(* IEC 61131-3 sources: Masterarbeit/sigmatek/lasalclass2/PW022_hardware/Class/_DriveMngBase (part 2) *)

    for x := 0 to SDDMAXENTRIES -1 do
      if (AxBuffer[x].pThis <> NIL) then
        if(AxBuffer[x].InitFinished = FALSE) & (AxBuffer[x].AxisOk = 1) then
          return;
        end_if;
      else
        exit;
      end_if;
    end_for;

    bdSettings.AxisInit := TRUE;

    if bVaranConnected then
      toVaran.ExternInitFinished();
    else
      MyPara.uiCmd := BUSIF_DRIVEMNGBASE_EXTERN_INIT_FINISH;
      ToBusIF.NewInst(#MyPara, #MyResult);
    end_if;

END_FUNCTION

FUNCTION _DriveMngBase::ResetAxisInit
  VAR
  	x       : USINT;
  END_VAR

    for x := 0 to SDDMAXENTRIES -1 do
      if (AxBuffer[x].pThis <> NIL) then
        if (AxBuffer[x].AxisOk = 1) then
          AxBuffer[x].InitFinished := FALSE;
        end_if;
      end_if;
    end_for;

END_FUNCTION

FUNCTION GLOBAL _DriveMngBase::CommunicationState
	VAR_OUTPUT
		retcode 	: DINT;
	END_VAR

  retcode := cOnline;

END_FUNCTION

FUNCTION _DriveMngBase::L2CmdFinished
	VAR_INPUT
		pPara 	: ^CmdStruct;
		pResult 	: ^results;
	END_VAR
	VAR_OUTPUT
		ret_code 	: iprStates;
	END_VAR

  ret_code := READY;

  L2Buffer[L2WrIndex].AxisNo := to_usint(pPara^.aPara[3]);
  L2Buffer[L2WrIndex].ParRW := to_usint(pPara^.aPara[1]);
  L2Buffer[L2WrIndex].ParNo := to_usint(pPara^.aPara[0]);
  L2Buffer[L2WrIndex].ParValue := pPara^.aPara[2];
  L2Buffer[L2WrIndex].bActive := TRUE;

  if pPara^.uiCmd = SDD_ASYNC_READY then
    L2Buffer[L2WrIndex].ParState := 0;
  else
    L2Buffer[L2WrIndex].ParState := 1;
    L2Buffer[L2WrIndex].ParError := to_sint(pPara^.aPara[4]);
  end_if;

  L2WrIndex += 1;
  L2NewEntry += 1;
  if L2WrIndex > (L2MAXINDEX - 1) then
    L2WrIndex := 0;
  end_if;

END_FUNCTION

FUNCTION VIRTUAL GLOBAL _DriveMngBase::CmdState::NewInst
	VAR_INPUT
		pPara 	: ^CmdStruct;
		pResult 	: ^results;
	END_VAR
	VAR_OUTPUT
		ret_code 	: iprStates;
	END_VAR
  VAR
    AxisNo          : USINT;
    ParRW           : USINT;
    ParNo           : USINT;
    retcode         : DINT;
    AxIndex         : USINT;
    RetcodeSizeLeft : UDINT;
    pActRetEntry    : ^_ParaRefreshBufEntry;
    i               : USINT;
    pThisRes        : ^UDINT;
    FoundAxis       : USINT;

    // Variables for CMD_GET_HARDWARE_DIAGNOSIS and CMD_GET_HARDWARE_TREE_ENTRY
    pStr_HWTRequested         : ^CHAR;
    us_HWTRequestedCurrIndex  : USINT;
    us_RequestedPlace         : USINT;
    us_RequestedAxis          : USINT;
    us_NextAxis               : USINT;
    us_NextPlace              : USINT;
    ud_StrSize                : UDINT;
    ud_TempSerNo              : UDINT;

    MyPara   : CmdStruct;
    MyResult : results;
  END_VAR

  pStr_HWTRequested         := NIL;
  us_HWTRequestedCurrIndex  := 0;
  us_RequestedPlace         := 16#FF;
  us_RequestedAxis          := 16#FF;
  us_NextAxis               := 16#FF;
  us_NextPlace              := 16#FF;
  ud_StrSize                := 0;
  ud_TempSerNo              := 0;

  ret_code := READY;

  CASE pPara^.uiCmd OF
  SDD_ASYNC_READY :

    // check the parameter number
    case (pPara^.aPara[0]) of

    SDD_I_HW :

      HWVersion := pPara^.aPara[2];
      DriveType := GetDriveType(pPara^.aPara[2]);
      bdWait4HwInfoResponse.I_HW := FALSE;

    SDD_I_TYPE :

      Parameter_I_Type := pPara^.aPara[2];
      bdWait4HwInfoResponse.I_Type := FALSE;

    SDD_I_SER :

      SerialNo := pPara^.aPara[2];
      bdWait4HwInfoResponse.I_SER := FALSE;

    SDD_I_FW :

      FwVersionInt :=  pPara^.aPara[2];
      bdWait4HwInfoResponse.I_FW := FALSE;
      SetFWVersion();

    SDD_I_BUILD :

      FWDateInt :=  pPara^.aPara[2]$UDINT;
      bdWait4HwInfoResponse.I_BUILD := FALSE;
      SetFwDate();

    else

      // Parameter for log file are dependent on the drive, usParaLogIdx is set in GetLogFileCyclic
      if pPara^.aPara[0] = s_LogFileV.usParaLogIdx then
        s_LogFileV.dParaLogValRd     := pPara^.aPara[2];
        s_LogFileV.bWait4LogFilePara := FALSE;
      end_if;

    end_case;

  SDD_ASYNC_ERROR :
    case pPara^.aPara[0] of

    SDD_I_HW :

      HWVersion := 16#7FFFFFFF;
      DriveType := _NotFound;
      bdWait4HwInfoResponse.I_HW := FALSE;

    SDD_I_TYPE :

      Parameter_I_Type := 16#7FFFFFFF;
      bdWait4HwInfoResponse.I_Type := FALSE;

    SDD_I_SER :

      SerialNo := 16#7FFFFFFF;
      bdWait4HwInfoResponse.I_SER := FALSE;

    SDD_I_FW :

      FwVersionInt :=  16#7FFFFFFF;
      bdWait4HwInfoResponse.I_FW := FALSE;

    SDD_I_BUILD :

      FWDateInt :=  16#7FFFFFFF;
      bdWait4HwInfoResponse.I_BUILD := FALSE;

    else

      // Parameter for log file are dependent on the drive, usParaLogIdx is set in GetLogFileCyclic
      if pPara^.aPara[0] = s_LogFileV.usParaLogIdx then
        s_LogFileV.dParaLogValRd     := 16#7FFFFFFF;
        s_LogFileV.bWait4LogFilePara := FALSE;
      end_if;

    end_case;

  SDD_GETVERSION :
    ret_code := READY;
    pResult^.uiLng := sizeof(UINT);
    pResult^.aData[0] := SDD_L2VERSION;
    pResult^.aData[1] := 0;

  SDD_ONLINEOK :

    ret_code := READY;
    pResult^.uiLng := sizeof(USINT);
    pResult^.aData[0] := to_usint(Online.read());

    // if the ringbuffer is allocated
    if ChangesRingBuffer.pStart then
      // we reset the ringbuffer which contains the changes
      ChangesRingBuffer.ActEntries := 0;
      ChangesRingBuffer.pWrite := ChangesRingBuffer.pRead := ChangesRingBuffer.pStart;
      _memset(ChangesRingBuffer.pStart, 16#00, SDDBUFFERENTRY*sizeof(_ParaRefreshBufEntry));
    end_if;

  SDD_RWPARLASAL2 :

    if Online.read() = 1 then
      ret_code := BUSY;

      // get Axisnumber
      AxisNo := to_usint(pPara^.aPara[0] AND 16#FF);

      // on SDD210 or SDD215 we fake the axis number of the 2nd axis for external use, so we have to correct it here
      if b_IsSDD21x & (AxisNo = 2) then // RamAnd 22.09.2010 16:12
        AxisNo := 3;
      end_if;

      AxIndex := GetAxIndex(AxisNo-1);

      if AxIndex = 16#FF then
        ret_code := ERROR;
        return;
      end_if;

      // read or write
      ParRw   := to_usint((pPara^.aPara[0] AND 16#FF00) SHR 8);
      // parameter number
      ParNo   := to_usint((pPara^.aPara[0] AND 16#FF0000) SHR 16);

      case ParRw of
      0 : // Read the parameter
        //if right I-HC code and scope buffer request then read 12 byte drive scope data over ID 0x2080 and SubID 0x09 is allowed
        if ((HWVersion and DRIVEMNG_DRIVESCOPE_SCOPE_BIT) = DRIVEMNG_DRIVESCOPE_SCOPE_BIT)
        & bLasalErrorBufferRequest = FALSE then

          case ParNo of
            251:
              AddASyncEntryDS402(AxisNo:=AxIndex, uiParaID:=DRIVEMNG_DRIVESCOPE_GETALL_PARAM, usParaSubID:=9, usRdWr:=0, pValue:=Nil, bsDataInfo:=2, pThisObj:= this, usEntry:=3);
              ret_code := Busy;

            252:
              //use always zero for SDD1X00 scope data
              pPara^.aPara[0] := (pPara^.aPara[0] AND (16#FFFFFF00)$DINT);
              ret_code := CmdState.GetState(pPara:=pPara, pResult:=pResult);

            253:
              //use always zero for SDD1X00 scope data
              pPara^.aPara[0] := (pPara^.aPara[0] AND (16#FFFFFF00)$DINT);
              ret_code := CmdState.GetState(pPara:=pPara, pResult:=pResult);

          else
            retcode := AddASyncEntry(AxisNo:= AxIndex, usParaNr:= ParNo , usRdWr:= ParRw, dValue:=0, pThisObj:= this, usEntry:=3);
          end_case;
        else
          retcode := AddASyncEntry(AxisNo:= AxIndex, usParaNr:= ParNo , usRdWr:= ParRw, dValue:=0, pThisObj:= this, usEntry:=3);
        end_if;

      1 : // Write the parameter
        //if right I-HC code then read 12 byte drive scope data over ID 0x2080 and SubID 0x09 is allowed
        if ((HWVersion and DRIVEMNG_DRIVESCOPE_SCOPE_BIT) = DRIVEMNG_DRIVESCOPE_SCOPE_BIT) then
          if ParNo = 249 then
            //remember which request come from Lasal2 (Drive Scope or Errorbuffer)
            if pPara^.aPara[1] > DRIVEMNG_DRIVESCOPE_SINDEX_RANGE then
              bLasalErrorBufferRequest := TRUE;
            else
              bLasalErrorBufferRequest := FALSE;
            end_if;
          end_if;
        end_if;

        retcode := AddASyncEntry(AxisNo:= AxIndex, usParaNr:= ParNo , usRdWr:= ParRw, dValue:=pPara^.aPara[1], pThisObj:= this, usEntry:=3);
      else
        ret_code := ERROR;
      end_case;

      if retcode < 0 then
        // internal failure
        Ret_code := ERROR;
      end_if;
    else
      ret_code := ERROR;
    end_if;

  SDD_GETAXISINUSE :
    ret_code := READY;
    pResult^.uiLng := sizeof(BDINT);
    pResult^.aData[0]$BDINT :=  AxIndizesL2;

  SDD_GETSERIE :
    retcode := READY;
    pResult^.uiLng := sizeof(USINT);
    if bVaranConnected then
      pResult^.aData[0] := toVaran.GetSeries();
    else
      //sdias drive connected
      MyPara.uiCmd  := BUSIF_DRIVEMNGBASE_SDD_GETSERIES;
      ToBusIF.NewInst(#MyPara, #MyResult);
      pResult^.aData[0] := MyResult.aData[0];
    end_if;

  // new commands in lasal communication version 4 (SDD_GET_CHANGE_CNT, SDD_GET_PARAMS)
  SDD_GET_CHANGE_CNT :
    retcode := READY;
    pResult^.uiLng := sizeof(UDINT);
    pResult^.aData[0]$^DINT := #ChangesRingBuffer.ActEntries;

  SDD_GET_PARAMS :
    retcode := READY;
    if ChangesRingBuffer.ActEntries then

      RetcodeSizeLeft := sizeof(pResult^.aData) - SIZEOF(UINT);
      pResult^.uiLng := 0;

      pActRetEntry := (#pResult^.aData[2])$^_ParaRefreshBufEntry;

      // as long as there are entries in change buffer and we still have some place in the return value array
      while ChangesRingBuffer.ActEntries & (RetcodeSizeLeft > sizeof(_ParaRefreshBufEntry)) do

        // store actual buffer entry in returncode
        pActRetEntry^ := ChangesRingBuffer.pRead^;

        // increase size of returncode in it's header
        pResult^.uiLng += sizeof(_ParaRefreshBufEntry);

        // decrease available size of returncode
        RetcodeSizeLeft -= sizeof(_ParaRefreshBufEntry);

        // increase pointer in retcode
        pActRetEntry += sizeof(_ParaRefreshBufEntry);

        // increase read pointer in ring buffer
        ChangesRingBuffer.pRead += sizeof(_ParaRefreshBufEntry);
        if ChangesRingBuffer.pRead >= ChangesRingBuffer.pEnd then
          ChangesRingBuffer.pRead := ChangesRingBuffer.pStart;
        end_if;

        // decrease available changes
        ChangesRingBuffer.ActEntries -= 1;
      end_while;

      // save number of entries in the first 2 byte of the array
      pResult^.aData[0]$UINT := pResult^.uiLng / sizeof(_ParaRefreshBufEntry);

      LastRetcode := pResult^;
    else
      // no changes to fetch
      pResult^.uiLng := 0;
    end_if;

  //++++++++++++++++++++++++++++++++++++++++++++++++++++++++++++++++++++++++++++++++++++++++++++++++++++++++++++++++++++
  SDD_GET_AXIS_PTR_LIST:

    ret_code := READY;

    //                    NoAxis    +  Thisptr per axis
    pResult^.uiLng := (sizeof(DINT) + AxCount * sizeof(UDINT))$UINT;

    // get no of axis
    pResult^.aData[0]$DINT := AxCount;

    // get this pointer of axis to resultbuffer (with increasing AxNumber)
    pThisRes := #pResult^.aData[4]$UDINT;
    FoundAxis := 0;
    for i := 0 to SDDMAXENTRIES-1 do
      AxIndex := GetAxIndexByAxisBit(1 SHL i);
      if AxIndex <> 16#FF then
        FoundAxis += 1;
        pThisRes^ := AxBuffer[AxIndex].pThis$UDINT;
        pThisRes += sizeof(UDINT);
      end_if;
      if FoundAxis = AxCount then
        // all avaliable found, exit loop
        exit;
      end_if;
    end_for;
    // fill space with NIL if a axis is not found
    while FoundAxis < AxCount do
      pThisRes^ := NIL;
      pThisRes += sizeof(UDINT);
      FoundAxis += 1;
    end_while;

  //++++++++++++++++++++++++++++++++++++++++++++++++++++++++++++++++++++++++++++++++++++++++++++++++++++++++++++++++++++
  CMD_GET_HARDWARE_DIAGNOSIS :

    pResult^.aData$t_HWCGetHardwareDiagnosisOut.retcode := _HWC_RETVAL_ERROR;
    ret_code := ERROR;

    pStr_HWTRequested := pPara^.aPara[0]$t_HWCGetHardwareDiagnosisIn.pStr_HardewareTreeEntry;

    // Check HWT String
    if pStr_HWTRequested then

      us_HWTRequestedCurrIndex := to_usint(pStr_HWTRequested$^UINT^ + 1); // +1 for 2byte length, points to end of HWT String

      if ( (pStr_HWTRequested + us_HWTRequestedCurrIndex - 1)^ = HWT_ESCAPE_DRIVE ) then // second to last byte is Drive escape sequence

        us_RequestedPlace := (pStr_HWTRequested + us_HWTRequestedCurrIndex)^; // Get passed place

        // Return State and Device ID and set retcode ----------------------------------------------------------
        pResult^.aData$t_HWCGetHardwareDiagnosisOut.ClassState := CmdState;

        pResult^.aData$t_HWCGetHardwareDiagnosisOut.ud_DeviceID := GetDrvDeviceID();

        if CmdState = _NoHardware then
          pResult^.aData$t_HWCGetHardwareDiagnosisOut.retcode := _HWC_RETVAL_ERROR_NO_HARDWARE;
        elsif CmdState = _WrongHardware then
          pResult^.aData$t_HWCGetHardwareDiagnosisOut.retcode := _HWC_RETVAL_ERROR_WRONG_HARDWARE;
        elsif CmdState = _NoCalibDataFound then
          pResult^.aData$t_HWCGetHardwareDiagnosisOut.retcode := _HWC_RETVAL_ERROR_NO_CALIB_DATA_FOUND;
        elsif CmdState <> _ClassOk then
          pResult^.aData$t_HWCGetHardwareDiagnosisOut.retcode := _HWC_RETVAL_ERROR_NO_HARDWARE;
        end_if;
        //------------------------------------------------------------------------------------------------------

        if CmdState= _ClassOk then

          // Search for Axis with the passed place
          for i := 0 to SDDMAXENTRIES - 1 do
            if AxBuffer[i].pThis then

              if ( AxBuffer[i].Place  = us_RequestedPlace ) then

                // Diagnosis info is stored with the axis class
                ret_code := AxBuffer[i].pThis$pVirtualBase^.NewInst(pPara, pResult);

                // FW Version ----------------------------------------------------------------------------------------------------------
                pResult^.aData[0]$t_HWCGetHardwareDiagnosisOut.pStr_FWVersion := #a_FWVersion[0];  // Will be overwritten if this pointer is not equal

                ud_StrSize := FwNumStr.GetLength() ;
                pResult^.aData[0]$t_HWCGetHardwareDiagnosisOut.pStr_FWVersion     := NIL;

                if ud_StrSize then

                  if (ud_StrSize < sizeof(a_FWVersion)) then // < to account for 0 termination
                    // Copy complete string
                    FwNumStr.GetDataAt(pData:=#a_FWVersion[0], udSize:=ud_StrSize, udAt:=0);
                    a_FWVersion[ud_StrSize] := 0; // 0 termination
                  else
                    // Copy part string
                    FwNumStr.GetDataAt(pData:=#a_FWVersion[0], udSize:=sizeof(a_FWVersion)-1, udAt:=0);
                    a_FWVersion[sizeof(a_FWVersion)-1] := 0; // 0 termination
                  end_if;

                  pResult^.aData[0]$t_HWCGetHardwareDiagnosisOut.pStr_FWVersion := #a_FWVersion[0];
                end_if;

                // HW Version
                pResult^.aData[0]$t_HWCGetHardwareDiagnosisOut.hd_HWVersion := HWVersion$UDINT;

                return;
              end_if;

            end_if;

          end_for;

          pResult^.aData$t_HWCGetHardwareDiagnosisOut.retcode := _HWC_RETVAL_ERROR_AXIS_MODULE_NOT_FOUND;
          ret_code := ERROR;

        end_if;

      elsif ( (pStr_HWTRequested + us_HWTRequestedCurrIndex - 1)^ = HWT_ESCAPE_AXIS ) &      // second to last byte is Axis escape sequence
            ( (pStr_HWTRequested + us_HWTRequestedCurrIndex - 3)^ = HWT_ESCAPE_DRIVE ) then

        us_RequestedPlace := (pStr_HWTRequested + us_HWTRequestedCurrIndex - 2)^; // Get passed place
        us_RequestedAxis  := (pStr_HWTRequested + us_HWTRequestedCurrIndex)^ + 1; // Get passed axisno (+1 AxisNo in HWT String run from 0 to 2)

        // Return State and Device ID and set retcode ----------------------------------------------------------
        pResult^.aData$t_HWCGetHardwareDiagnosisOut.ClassState := CmdState;

        pResult^.aData$t_HWCGetHardwareDiagnosisOut.ud_DeviceID := GetDrvDeviceID();

        if CmdState = _NoHardware then
          pResult^.aData$t_HWCGetHardwareDiagnosisOut.retcode := _HWC_RETVAL_ERROR_NO_HARDWARE;
        elsif CmdState = _WrongHardware then
          pResult^.aData$t_HWCGetHardwareDiagnosisOut.retcode := _HWC_RETVAL_ERROR_WRONG_HARDWARE;
        elsif CmdState = _NoCalibDataFound then
          pResult^.aData$t_HWCGetHardwareDiagnosisOut.retcode := _HWC_RETVAL_ERROR_NO_CALIB_DATA_FOUND;
        elsif CmdState <> _ClassOk then
          pResult^.aData$t_HWCGetHardwareDiagnosisOut.retcode := _HWC_RETVAL_ERROR_NO_HARDWARE;
        end_if;
        //------------------------------------------------------------------------------------------------------

        if CmdState= _ClassOk then

          // Search for Axis with the passed place and axisno
          for i := 0 to SDDMAXENTRIES - 1 do
            if AxBuffer[i].pThis then

              if ( AxBuffer[i].Place  = us_RequestedPlace ) &
                 ( AxBuffer[i].AxisNo = us_RequestedAxis  ) then

                ret_code := AxBuffer[i].pThis$pVirtualBase^.NewInst(pPara, pResult);
                return;
              end_if;

            end_if;

          end_for;

          pResult^.aData$t_HWCGetHardwareDiagnosisOut.retcode := _HWC_RETVAL_ERROR_AXIS_MODULE_NOT_FOUND;
          ret_code := ERROR;

        end_if;
      else

        // Return diagnosis for the DriveMng

        // Return State and Device ID and set retcode ----------------------------------------------------------
        pResult^.aData$t_HWCGetHardwareDiagnosisOut.ClassState := CmdState;

        pResult^.aData$t_HWCGetHardwareDiagnosisOut.ud_DeviceID := GetBusDeviceID();

        if CmdState = _NoHardware then
          pResult^.aData$t_HWCGetHardwareDiagnosisOut.retcode := _HWC_RETVAL_ERROR_NO_HARDWARE;
        elsif CmdState = _WrongHardware then
          pResult^.aData$t_HWCGetHardwareDiagnosisOut.retcode := _HWC_RETVAL_ERROR_WRONG_HARDWARE;
        elsif CmdState = _NoCalibDataFound then
          pResult^.aData$t_HWCGetHardwareDiagnosisOut.retcode := _HWC_RETVAL_ERROR_NO_CALIB_DATA_FOUND;
        elsif CmdState <> _ClassOk then
          pResult^.aData$t_HWCGetHardwareDiagnosisOut.retcode := _HWC_RETVAL_ERROR_NO_HARDWARE;
        end_if;
        //------------------------------------------------------------------------------------------------------

        if CmdState= _ClassOk then

          //Data which is already in HWK available
          pResult^.aData[0]$t_HWCGetHardwareDiagnosisOut.ud_DeviceID := DeviceID;
          pResult^.aData[0]$t_HWCGetHardwareDiagnosisOut.ud_VendorID := VendorID;

          pResult^.aData$t_HWCGetHardwareDiagnosisOut.retcode := _HWC_RETVAL_OK;
          ret_code := READY;

        end_if;
      end_if;

    end_if;

  //++++++++++++++++++++++++++++++++++++++++++++++++++++++++++++++++++++++++++++++++++++++++++++++++++++++++++++++++++++
  CMD_GET_HARDWARE_TREE_ENTRY:

    ret_code := ERROR;
    pResult^.aData[0]$t_HWCGetHardwareTreeEntryOut.retcode := _HWC_RETVAL_ERROR;

    pStr_HWTRequested := pPara^.aPara[0]$t_HWCGetHardwareTreeEntryIn.pStr_LastHardewareTreeEntry;

    if pStr_HWTRequested then

      us_HWTRequestedCurrIndex := to_usint(pStr_HWTRequested$^UINT^ + 1); // +1 for 2byte length, points to end of HWT String

      // -----------------------------------------------------------------------------------------------------------------------------
      // Return 1st axis at place, if no axis at place return next place
      if ( (pStr_HWTRequested + us_HWTRequestedCurrIndex - 1)^ = HWT_ESCAPE_DRIVE ) then

        us_RequestedPlace := (pStr_HWTRequested + us_HWTRequestedCurrIndex)^; // Get last place

        // Find 1.st axis at place
        us_NextAxis := 16#FF;

        for i := 0 to SDDMAXENTRIES - 1 do

          if (AxBuffer[i].pThis) &
             (AxBuffer[i].Place = us_RequestedPlace) &
             (AxBuffer[i].AxisNo < us_NextAxis) then

            us_NextAxis := to_usint(AxBuffer[i].AxisNo);
          end_if;

        end_for;

        if (us_NextAxis < 16#FF) then
          // Copy string and add axis no
          // Copy passed string
          _memcpy(ptr1 := #a_HWTEntryStr[0]
                , ptr2 := pStr_HWTRequested
                , cntr := pStr_HWTRequested^$UINT+2); // +2 for 2 byte length

          // Add Escape Sequence axis
          a_HWTEntryStr[0]$UINT += 1;
          a_HWTEntryStr[a_HWTEntryStr[0]$UINT+1] := HWT_ESCAPE_AXIS;

          // Add axis no
          a_HWTEntryStr[0]$UINT += 1;
          a_HWTEntryStr[a_HWTEntryStr[0]$UINT+1] := us_NextAxis - 1; // -1 AxisNo in HWT String run from 0 to 2

          // Set return pointer
          pResult^.aData[0]$t_HWCGetHardwareTreeEntryOut.pStr_NextHardewareTreeEntry := #a_HWTEntryStr[0];

          ret_code := READY;
          pResult^.aData[0]$t_HWCGetHardwareTreeEntryOut.retcode := _HWC_RETVAL_OK_HWTSTR_RETURNED;

          return;
        else

          // Find min next place
          us_NextPlace := 16#FF;

          // No Axis found at this place, return next place
          for i := 0 to SDDMAXENTRIES - 1 do

            if (AxBuffer[i].Place > us_RequestedPlace) &  // Next Place must be the minmum place that is greater then the passed palce
               (AxBuffer[i].Place < us_NextPlace) then

              us_NextPlace := to_usint(AxBuffer[i].Place);
            end_if;

          end_for;

          if (us_NextPlace < 16#FF) then
            // Copy string and replace place
            // Copy passed string
            _memcpy(ptr1 := #a_HWTEntryStr[0]
                  , ptr2 := pStr_HWTRequested
                  , cntr := pStr_HWTRequested^$UINT+2); // +2 for 2 byte length

            // replace place
            a_HWTEntryStr[a_HWTEntryStr[0]$UINT+1] := us_NextPlace;

            // Set return pointer
            pResult^.aData[0]$t_HWCGetHardwareTreeEntryOut.pStr_NextHardewareTreeEntry := #a_HWTEntryStr[0];

            ret_code := READY;
            pResult^.aData[0]$t_HWCGetHardwareTreeEntryOut.retcode := _HWC_RETVAL_OK_HWTSTR_RETURNED;
            return;

          else

            ret_code := READY;
            pResult^.aData[0]$t_HWCGetHardwareTreeEntryOut.retcode := _HWC_RETVAL_OK_END_OF_LIST;
            return;
          end_if;

        end_if;

      // -----------------------------------------------------------------------------------------------------------------------------
      // return next axis, if last axis at passed place return next place
      elsif ( (pStr_HWTRequested + us_HWTRequestedCurrIndex - 1)^ = HWT_ESCAPE_AXIS )  &
            ( (pStr_HWTRequested + us_HWTRequestedCurrIndex - 3)^ = HWT_ESCAPE_DRIVE ) then  // Must be 1st entry second to last byte is next Axis escape sequence

        us_RequestedPlace := (pStr_HWTRequested + us_HWTRequestedCurrIndex - 2)^; // Get last place
        us_RequestedAxis  := (pStr_HWTRequested + us_HWTRequestedCurrIndex)^ + 1; // Get last axisno (+1 AxisNo in HWT String run from 0 to 2)

        // Find min next axis
        us_NextAxis := 16#FF;

        for i := 0 to SDDMAXENTRIES - 1 do

          if (AxBuffer[i].pThis) &
             (AxBuffer[i].Place = us_RequestedPlace) &
             (AxBuffer[i].AxisNo > us_RequestedAxis) &
             (AxBuffer[i].AxisNo < us_NextAxis) then

            us_NextAxis := to_usint(AxBuffer[i].AxisNo);
          end_if;

        end_for;

        if (us_NextAxis < 16#FF) then

          // Copy string and replace AxisNo
          // Copy passed string
          _memcpy(ptr1 := #a_HWTEntryStr[0]
                , ptr2 := pStr_HWTRequested
                , cntr := pStr_HWTRequested^$UINT+2); // +2 for 2 byte length

          // replace AxisNo
          a_HWTEntryStr[a_HWTEntryStr[0]$UINT+1] := us_NextAxis - 1;  // -1 AxisNo in HWT String run from 0 to 2

          // Set return pointer
          pResult^.aData[0]$t_HWCGetHardwareTreeEntryOut.pStr_NextHardewareTreeEntry := #a_HWTEntryStr[0];

          ret_code := READY;
          pResult^.aData[0]$t_HWCGetHardwareTreeEntryOut.retcode := _HWC_RETVAL_OK_HWTSTR_RETURNED;
          return;

        else

          // Find min next place
          us_NextPlace := 16#FF;

          // Search for next Place
          for i := 0 to SDDMAXENTRIES - 1 do

            if (AxBuffer[i].pThis) &
               (AxBuffer[i].Place > us_RequestedPlace) &
               (AxBuffer[i].Place < us_NextPlace) then

              us_NextPlace := to_usint(AxBuffer[i].Place);
            end_if;
          end_for;

          if (us_NextPlace < 16#FF) then

            // Copy string and replace place
            // Copy passed string
            _memcpy(ptr1 := #a_HWTEntryStr[0]
                  , ptr2 := pStr_HWTRequested
                  , cntr := pStr_HWTRequested^$UINT+2); // +2 for 2 byte length

            // Throw away axis info
            a_HWTEntryStr[0]$UINT -= 2;

            // replace place
            a_HWTEntryStr[a_HWTEntryStr[0]$UINT+1] := us_NextPlace;

            // Set return pointer
            pResult^.aData[0]$t_HWCGetHardwareTreeEntryOut.pStr_NextHardewareTreeEntry := #a_HWTEntryStr[0];

            ret_code := READY;
            pResult^.aData[0]$t_HWCGetHardwareTreeEntryOut.retcode := _HWC_RETVAL_OK_HWTSTR_RETURNED;
            return;
          else

            ret_code := READY;
            pResult^.aData[0]$t_HWCGetHardwareTreeEntryOut.retcode := _HWC_RETVAL_OK_END_OF_LIST;
            return;

          end_if;

        end_if;

      // -----------------------------------------------------------------------------------------------------------------------------
      else  // 1st call after manager, find and return min valid place

        // Find min next place
        us_NextPlace := 16#FF;

        // Search for next Place
        for i := 0 to SDDMAXENTRIES - 1 do

          if (AxBuffer[i].pThis) &
             (AxBuffer[i].Place < us_NextPlace) then

            us_NextPlace := to_usint(AxBuffer[i].Place);
          end_if;
        end_for;

        if (us_NextPlace < 16#FF) then
          // Copy 1st part of HWT
          _memcpy(ptr1 := #a_HWTEntryStr[0]
                , ptr2 := pStr_HWTRequested
                , cntr := pStr_HWTRequested^$UINT+2); // +2 for 2 byte length

          // Add Escape Sequence drive
          a_HWTEntryStr[0]$UINT += 1;
          a_HWTEntryStr[a_HWTEntryStr[0]$UINT+1] := HWT_ESCAPE_DRIVE;

          // Add Place
          a_HWTEntryStr[0]$UINT += 1;
          a_HWTEntryStr[a_HWTEntryStr[0]$UINT+1] := us_NextPlace;

          // Set return pointer
          pResult^.aData[0]$t_HWCGetHardwareTreeEntryOut.pStr_NextHardewareTreeEntry := #a_HWTEntryStr[0];

          ret_code := READY;
          pResult^.aData[0]$t_HWCGetHardwareTreeEntryOut.retcode := _HWC_RETVAL_OK_HWTSTR_RETURNED;
          return;
        else

          ret_code := READY;
          pResult^.aData[0]$t_HWCGetHardwareTreeEntryOut.retcode := _HWC_RETVAL_OK_END_OF_LIST;
          return;

        end_if;

      end_if;

//    else
//
//      // Error, Need valid HWT String from Manager
//      return;
    end_if;

  //*******************************************************************************************************************
  SDD_GET_DEVICESERIALNO:
    ret_code := READY;
    //Get Serial No. of Head of MDD100
    //Here: Get Serial No of all devices (also of VAC)
    if bVaranConnected then
      pResult^.uiLng := 1 + (toVaran.SerialNoStr.GetLength())$UINT;
      toVaran.SerialNoStr.GetDataAt(#pResult^.aData[0], pResult^.uiLng, 0);
    end_if;

  //*******************************************************************************************************************
  SDD_GET_MNG_TRANSPARENT:
    ret_code := READY;
   //Get transparent information from VaranCommunication object. used to not show transparent objects in DiasDriveOnline Window
    pResult^.uiLng := sizeof(DINT);
    if bVaranConnected then
      pResult^.aData[0]$DINT := toVaran.Transparent.Read();
    else
      pResult^.aData[0]$DINT := 0$DINT;
    end_if;

  //*******************************************************************************************************************
  SDD_GETFILE: //command will be called from application

    ret_code := ERROR;

    //Check version 1
    if pPara^.aPara[0] = SDD_GETFILE_VER_1 then
      //Call method
      ret_code := GetFile(pDestinationDPNE := pPara^.aPara[1]$^CHAR
                        , pFileNameDrive   := pPara^.aPara[2]$^CHAR
                        , pFilePathDrive   := pPara^.aPara[3]$^CHAR
                        , pdError          := pPara^.aPara[4]$^DINT
                        );
    elsif pPara^.aPara[4] then
      (pPara^.aPara[4]$^DINT)^ := DRIVEMNG_FILE_HANDLING_RETCODE_CMDVERSION_NOTSUPPORTED;
    end_if;

    pResult^.uiLng := 4;
    pResult^.aData[0]$DINT := SDD_GETFILE_VER_MAX;  //max supported version

  //*******************************************************************************************************************
  SDD_GETLOGFILE: //command will be called from application

    ret_code := ERROR; //unsupported version

    //Check version 1
    if pPara^.aPara[0] = SDD_GETLOGFILE_VER_1 then
      //Call method
      ret_code := GetLogFile(pDestinationDPNE  := pPara^.aPara[1]$^CHAR
                           , pdError           := pPara^.aPara[2]$^DINT
                           );
    //Check version 2
    elsif pPara^.aPara[0] = SDD_GETLOGFILE_VER_2 then
      //Call method
      ret_code := GetLogFile(pDestinationDPNE  := pPara^.aPara[1]$^CHAR
                           , pdError           := pPara^.aPara[2]$^DINT
                           , udFileSelectID    := pPara^.aPara[3]$UDINT
                           );
    elsif pPara^.aPara[2] then
      (pPara^.aPara[2]$^DINT)^ := DRIVEMNG_FILE_HANDLING_RETCODE_CMDVERSION_NOTSUPPORTED;
    end_if;

    pResult^.uiLng := 4;
    pResult^.aData[0]$DINT := SDD_GETLOGFILE_VER_MAX;  //max supported version

  //*******************************************************************************************************************
  SDD_GETFILESTATE:  //command will be called from application

    ret_code := ERROR; //unsupported version

    //Check version 1
    if pPara^.aPara[0] = SDD_GETFILESTATE_VER_1 then
      //Call method
      ret_code := GetFileState(pdError      :=  pPara^.aPara[1]$^DINT
                             , pdProgress   :=  pPara^.aPara[2]$^DINT
                             , pudBytesRead :=  pPara^.aPara[3]$^UDINT
                              );
    elsif pPara^.aPara[1] then
      (pPara^.aPara[1]$^DINT)^ := DRIVEMNG_FILE_HANDLING_RETCODE_CMDVERSION_NOTSUPPORTED;
    end_if;

    pResult^.uiLng := 4;
    pResult^.aData[0]$DINT := SDD_GETFILESTATE_VER_MAX;  //max supported version

  //*******************************************************************************************************************
  SDD_SETFILE: //command will be called from application

    ret_code := ERROR;

    //Check version 1
    if pPara^.aPara[0] = SDD_SETFILE_VER_1 then
      //Call method
      ret_code := SetFile(pWriteData      :=  pPara^.aPara[1]$^void
                        , udWriteDataLen  :=  pPara^.aPara[2]$UDINT
                        , pFilePathDrive  :=  pPara^.aPara[3]$^cHAR
                        , pFileNameDrive  :=  pPara^.aPara[4]$^cHAR
                        , pdError         :=  pPara^.aPara[5]$^DINT
                        );
    elsif pPara^.aPara[5] then
      (pPara^.aPara[5]$^DINT)^ := DRIVEMNG_FILE_HANDLING_RETCODE_CMDVERSION_NOTSUPPORTED;
    end_if;

    pResult^.uiLng := 4;
    pResult^.aData[0]$DINT := SDD_SETFILE_VER_MAX;  //max supported version

//*******************************************************************************************************************
  SDD_GETFILESIZE:  //command will be called from application

    ret_code := ERROR; //unsupported version

    //Check version 1
    if pPara^.aPara[0] = SDD_GETFILESIZE_VER_1 then
      //Call method
      ret_code := GetFileSize(pFileNameDrive  :=  pPara^.aPara[1]$^CHAR
                            , pFilePathDrive  :=  pPara^.aPara[2]$^CHAR
                            , pudSize         :=  pPara^.aPara[3]$^UDINT
                            , pdError         :=  pPara^.aPara[4]$^DINT
                            );
    elsif pPara^.aPara[4] then
      (pPara^.aPara[4]$^DINT)^ := DRIVEMNG_FILE_HANDLING_RETCODE_CMDVERSION_NOTSUPPORTED;
    end_if;

    pResult^.uiLng := 4;
    pResult^.aData[0]$DINT := SDD_GETFILESIZE_VER_MAX;  //max supported version

//*******************************************************************************************************************
  SDD_GETFILEBUFFER:  //command will be called from application

    ret_code := ERROR; //unsupported version

    //Check version 1
    if pPara^.aPara[0] = SDD_GETFILEBUFFER_VER_1 then
      //Call method

      ret_code := GetFileBuffer(pFileNameDrive  :=  pPara^.aPara[1]$^CHAR
                              , pFilePathDrive  :=  pPara^.aPara[2]$^CHAR
                              , udBufferSize    :=  pPara^.aPara[3]$UDINT
                              , pDataBuffer     :=  pPara^.aPara[4]$^void
                              , udDataLenToRead :=  pPara^.aPara[5]$UDINT
                              , pdError         :=  pPara^.aPara[6]$^DINT
                              );
    elsif pPara^.aPara[6] then
      (pPara^.aPara[6]$^DINT)^ := DRIVEMNG_FILE_HANDLING_RETCODE_CMDVERSION_NOTSUPPORTED;
    end_if;

    pResult^.uiLng := 4;
    pResult^.aData[0]$DINT := SDD_GETFILEBUFFER_VER_MAX;  //max supported version

  end_case;

END_FUNCTION

FUNCTION VIRTUAL GLOBAL _DriveMngBase::CmdState::GetState
	VAR_INPUT
		pPara 	: ^CmdStruct;
		pResult 	: ^results;
	END_VAR
	VAR_OUTPUT
		ret_code 	: iprStates;
	END_VAR
  VAR
  	x         : BOOL;
    IntRdIndex  : DINT;
    AxisNo      : USINT;
    ParRW       : USINT;
    ParNo       : USINT;
  END_VAR

  ret_code := READY;

  case pPara^.uiCmd of

  SDD_RWPARLASAL2 :

    ret_code := BUSY;

    // get Axisnumber
    AxisNo := to_usint(pPara^.aPara[0] AND 16#FF) - 1;

    // on SDD210 or SDD215 we fake the axis number of the 2nd axis for external use, so we have to correct it here
    if b_IsSDD21x & (AxisNo = 1) then // RamAnd 22.09.2010 16:12
      AxisNo := 2;
    end_if;

    // read or write
    ParRw   := to_usint((pPara^.aPara[0] AND 16#FF00) SHR 8);
    // parameter number
    ParNo   := to_usint((pPara^.aPara[0] AND 16#FF0000) SHR 16);

    x := FALSE;
    if L2NewEntry <> 0 then
      for IntRdIndex := 0 to (L2MAXINDEX - 1) do
        // now check if the right command is available
        if ((AxisNo =  L2Buffer[IntRdIndex].AxisNo) | (AxisNo = 0xFF)) & //0xFF for drive scope parameter and SDD1X00 drives
           ParRw = L2Buffer[IntRdIndex].ParRW &
           ParNo = L2Buffer[IntRdIndex].ParNo  &
           L2Buffer[IntRdIndex].bActive = TRUE then
           // we found the correct info
           pResult^.uiLng := 8; // Result info hat 8 Byte
           pResult^.aData[0] := AxisNo;
           pResult^.aData[1] := L2Buffer[IntRdIndex].ParState ;// hier steht ob ein Error vorhanden ist oder Nicht
           if L2Buffer[IntRdIndex].ParState = 0 then
            pResult^.aData[2] := ParRw;
           else
            pResult^.aData[2] := to_usint(L2Buffer[IntRdIndex].ParError);
           end_if;
           pResult^.aData[3] := ParNo;
           pResult^.aData[4]$DINT := L2Buffer[IntRdIndex].ParValue;

           ret_code := READY;

           // Daten werden gelöscht :
           L2Buffer[IntRdIndex].AxisNo := 0;
           L2Buffer[IntRdIndex].bActive := FALSE;
           L2NewEntry -= 1;
           if L2NewEntry < 0 then
            L2NewEntry := 0;
           end_if;
           exit;
        end_if;
      end_for;

    end_if;

  else
    ret_code := NewInst(pPara, pResult);
  end_case;

END_FUNCTION

FUNCTION GLOBAL _DriveMngBase::GetAxisWrPtr
	VAR_INPUT
		usAxis 	: USINT;
	END_VAR
	VAR_OUTPUT
		ptr 	: ^_VaranDriveBase::t_WriteValuePtr;
	END_VAR
  VAR
    MyPara   : CmdStruct;
    MyResult : results;
  END_VAR

  if usAxis >= 0 & usAxis < SDDMAXENTRIES then //HasHan
    if bVaranConnected then
      ptr := toVaran.GetAxisWrPtr(AxisNr:=AxBuffer[usAxis].AxisIndex);
    else
      MyPara.uiCmd    := BUSIF_DRIVEMNGBASE_GET_AXIS_WR_PTR;
      MyPara.aPara[0] := to_dint(AxBuffer[usAxis].AxisIndex);
      ToBusIF.NewInst(#MyPara, #MyResult);
      ptr := MyResult.aData[0]$^_VaranDriveBase::t_WriteValuePtr;
    end_if;
  end_if;

END_FUNCTION

FUNCTION GLOBAL _DriveMngBase::GetAxisRdPtr
	VAR_INPUT
		usAxis 	: USINT;
	END_VAR
	VAR_OUTPUT
		ptr 	: ^_VaranDriveBase::t_ReadValuePtr;
	END_VAR
  VAR
    MyPara   : CmdStruct;
    MyResult : results;
  END_VAR

  if usAxis >= 0 & usAxis < SDDMAXENTRIES then //HasHan
    if bVaranConnected then
      ptr := toVaran.GetAxisRdPtr(AxisNr:=AxBuffer[usAxis].AxisIndex);
    else
      MyPara.uiCmd    := BUSIF_DRIVEMNGBASE_GET_AXIS_RD_PTR;
      MyPara.aPara[0] := to_dint(AxBuffer[usAxis].AxisIndex);
      ToBusIF.NewInst(#MyPara, #MyResult);
      ptr := MyResult.aData[0]$^_VaranDriveBase::t_ReadValuePtr;
    end_if;
  end_if;

END_FUNCTION

FUNCTION GLOBAL _DriveMngBase::InitDrive
	VAR_INPUT
		Mode 	: USINT;
	END_VAR
  VAR
    UserPara     : CmdStruct;
    UserResult   : Results;
    x            : USINT;
    pThisNewInst : ^void;
  END_VAR

  if bVaranConnected then
    toVaran.InitDrive();
  else
    UserPara.uiCmd := BUSIF_DRIVEMNGBASE_INIT_DRIVE;
    ToBusIF.NewInst(#UserPara, #UserResult);
  end_if;

  for x := 0 to (SDDMAXENTRIES - 1) do
    if (AxBuffer[x].pThis <> NIL) then
      if (AxBuffer[x].AxisOk = 1) then
        if Mode = 0 then
          UserPara.uiCmd := SDD_INITAXLE;
        else
          UserPara.uiCmd := SDD_URINITAXLE;
        end_if;

        pThisNewInst := AxBuffer[x].pThis;
        pThisNewInst$^VirtualBase^.NewInst(#UserPara, #UserResult);
      end_if;
    end_if;
  end_for;

END_FUNCTION

FUNCTION _DriveMngBase::GetAxIndex
	VAR_INPUT
		AxisNo 	: USINT;
	END_VAR
	VAR_OUTPUT
		AxIndex 	: USINT;
	END_VAR
  VAR
  	x     : USINT;
  END_VAR

  AxIndex := 16#FF;

  for x := 0 to (SDDMAXENTRIES - 1) do
    if (AxBuffer[x].pThis <> NIL) then
      if (AxBuffer[x].AxisOk = 1) & (AxBuffer[x].AxisIndex = AxisNo) then
        AxIndex := x;
        exit;
      end_if;
    else
      exit;
    end_if;
  end_for;

END_FUNCTION

FUNCTION _DriveMngBase::GetAxIndexByAxisBit
	VAR_INPUT
		AxisBit 	: BDINT;
	END_VAR
	VAR_OUTPUT
		AxIndex 	: USINT;
	END_VAR
  VAR
  	x     : USINT;
  END_VAR

  AxIndex := 16#FF;

  for x := 0 to (SDDMAXENTRIES - 1) do
    if (AxBuffer[x].pThis <> NIL) then
      if (AxBuffer[x].AxisBit = AxisBit) then
        AxIndex := x;
        exit;
      end_if;
    else
      exit;
    end_if;
  end_for;

END_FUNCTION

FUNCTION _DriveMngBase::GetFirstAxIndex
	VAR_OUTPUT
		AxIndex 	: USINT;
	END_VAR
  VAR
  	x     : USINT;
  END_VAR

  AxIndex := 16#FF;

  for x := 0 to (SDDMAXENTRIES - 1) do
    if (AxBuffer[x].pThis <> NIL) then
      if (AxBuffer[x].AxisOk = 1) then
        AxIndex := x;
        exit;
      end_if;
    else
      exit;
    end_if;
  end_for;

END_FUNCTION

FUNCTION _DriveMngBase::SetFwVersion
VAR
  szValue     : ARRAY[0..19] of CHAR;
  StrLen      : UDINT;
END_VAR

  Bin2Ascii(pt:=#szValue[0], value:=FwVersionInt, format:=16#820);
  StrLen := _strlen(#szValue[0]);
  FwNumStr.WriteDataOff(udLen:= Strlen, udOff:=0, pData:= #szValue[0]);

END_FUNCTION

FUNCTION _DriveMngBase::SetFwDate
VAR
	szValue     : ARRAY[0..19] of CHAR;
  szFwDate    : ARRAY[0..99] of CHAR;
  StrLen      : UDINT;
  Value       : UDINT;
  tmpYear     : UDINT;
END_VAR

  // Ermitteln des Tages
  Value := FWDateInt AND 16#003F0000;
  Value := Value SHR 16;
  Bin2Ascii(pt:=#szValue[0], value:=Value$DINT, format:=16#102);
  _strcpy(#szFwDate[0], #szValue[0]);
  _strcat(#szFwDate[0], ".");

  // ermitteln des Monats
  Value := FWDateInt AND 16#0F000000;
  Value := Value SHR 24;
  Bin2Ascii(pt:=#szValue[0], value:=Value$DINT, format:=16#102);
  _strcat(#szFwDate[0], #szValue[0]);
  _strcat(#szFwDate[0], ".");

  // ermitteln des Jahres
  Value := FWDateInt AND 16#F0000000;
  Value := Value SHR 28;

  //Newer firmwares >= 2016 are using 2 Bits more, which where originally reserved for day, to have more bits to display year dates.
  //With this change we can display year dates until 2063 instead of 2015,
  tmpYear := FWDateInt AND 16#00C00000;
  tmpYear := tmpYear SHR 18; //Shift Right 18 instead of 22 because these two bits are bit 4 and 5 for the year
  Value := Value OR tmpYear;

  Value += 2000;
  Bin2Ascii(pt:=#szValue[0], value:=Value$DINT, format:=16#800);
  _strcat(#szFwDate[0], #szValue[0]);
  _strcat(#szFwDate[0], " ");

  // ermitteln der Stunde
  Value := FWDateInt AND 16#0000FF00;
  Value := Value SHR 8;
  Bin2Ascii(pt:=#szValue[0], value:=Value$DINT, format:=16#102);
  _strcat(#szFwDate[0], #szValue[0]);
  _strcat(#szFwDate[0], ":");

  // ermitteln der Minuten
  Value := FWDateInt AND 16#000000FF;
  Bin2Ascii(pt:=#szValue[0], value:=Value$DINT, format:=16#102);
  _strcat(#szFwDate[0], #szValue[0]);

  StrLen := _strlen(#szFwDate[0]);
  FwDatetr.WriteDataOff(udLen:= Strlen, udOff:=0, pData:= #szFwDate[0]);

END_FUNCTION

(*
Der String kann folgendermaßen formatiert werden.
xxxx 0000 0000 0000     xxxx = keine Funktion.
     .... .... ****     Anzahl der Dezimalstellen.
     .... **** ....     Position des Dezimalpunkts.
     ...* .... ....     Vornullen (Anzahl der Dezimalstellen).
     ..*. .... ....     Nachkomma Nullen.
     .*.. .... ....     Vorzeichen unmittelbar vor wert (-3 ansonsten - 3).
     *... .... ....     Anzahl der Stellen automatisch ermitteln.

*)

FUNCTION _DriveMngBase::Bin2Ascii
	VAR_INPUT
		pt 	: ^CHAR;
		value 	: DINT;
		format 	: BINT;
	END_VAR
  VAR
    tmp    : DINT;
    nk     : UINT;
    dig    : UINT;
    hp     : ^CHAR;
    pd     : UINT;
    h      : UINT;
  END_VAR

  if((format AND 16#000F) = 0) then
    format := format OR 16#0800;
  end_if;

  if(format AND 16#0800) then
    tmp  := value;
    if tmp = 0 then
      dig := 1;
    else
      dig := 0;
    end_if;

    while(tmp) do

      tmp := tmp / 10;
      dig += 1;
    end_while;

    nk := ((format SHR 4) AND 16#0F);

    if(nk >= dig) then
      dig := nk + 1;
    end_if;

    format := (format AND 16#FFF0) OR (dig AND 16#000F);
  end_if;

  dig := (format and 16#0F);        // Anzahl der Stellen
  hp  := pt + dig;                  // pointer auf String-Ende
  tmp := value;                     // Zahl
  pd  := (format shr 4) and 16#0F;  // position des Komma

  if(value < 0) then    // kontrolle ob Zahl negativ
    hp    += 1;
    value := -value;    // Zahl * (-1)
    pt^   := '-';       // Erstes Zeichen auf '-' setzen
  end_if;

  if(format and 16#0200) then // Nachnullen löschen
    h := pd;
    while(h) do               // Nur Nullen hinter Komma
      h -= 1;
      if((value mod 10) = 0) then // Ist Ziffer Null?
        value := value / 10;      // wenn ja, Null löschen
        pd -= 1;
      else
        h := 0;
      end_if;

    end_while;
  end_if;

  if(pd <> 0) then       // Komma noch zu setzen?
    hp += 1;
  end_if;

  hp^ := 0;               // String mit Ascii-0 abschließen
  hp  -= 1;

  repeat
    hp^   := '0' + TO_USINT(value mod 10);  //akt. Ziffer
    hp    -= 1;
    pd    -= 1;
    dig   -= 1;
    if(pd = 0)then    // Komma setzen?
      hp^ := '.';
      hp -= 1;
    end_if;

    value := value / 10;   // nächste Ziffer

    if((dig = 0) & (value <> 0)) then // Zahl zu groß
      pt^   := '?';   // Formatfehler
      value := 0;
    end_if;
  until(value = 0) end_repeat;

  if(dig > 0) then  // mit Vornullen auffüllen
    repeat          // so lange bis Digits auf Null
      if((format and 16#0100)|(pd$INT >= 0)) then   // Vornullen im
        hp^ := '0';   // Format angegeben?
      else            // formatfehler (digit zu groß und keine Vornullen)
        pt^   := '?'; // Formatfehler
        value := 0;
      end_if;
      pd -= 1;
      hp -= 1;
      if(pd = 0) then // Komma setzen
        hp^ := '.';
        hp -= 1;
      end_if;
      dig -= 1;
    until(dig = 0) end_repeat;  // letzte Ziffer?
  end_if;

END_FUNCTION

FUNCTION VIRTUAL GLOBAL _DriveMngBase::RetryCounter::Read
	VAR_OUTPUT
		output (EAX) 	: UDINT;
	END_VAR
  VAR
    MyPara   : CmdStruct;
    MyResult : results;
  END_VAR

  if bVaranConnected then
    RetryCounter := toVaran.RetryCounter.Read();
  else
    MyPara.uiCmd  := BUSIF_DRIVEMNGBASE_READ_RETRY_COUNTER;
    ToBusIF.NewInst(#MyPara, #MyResult);
    RetryCounter := MyResult.aData[0]$UDINT;
  end_if;

  output := RetryCounter;

END_FUNCTION

FUNCTION GLOBAL _DriveMngBase::SetSyncEntry
	VAR_INPUT
		usAxis 	: USINT;
		usValue 	: USINT;
		usPData 	: DINT;
	END_VAR
	VAR_OUTPUT
		retcode 	: DINT;
	END_VAR
  VAR
    MyPara   : CmdStruct;
    MyResult : results;
  END_VAR

  if usAxis >= 0 & usAxis < SDDMAXENTRIES then //HasHan
    if bVaranConnected then
      retcode:=toVaran.SetSyncParameter(us_Axis:=AxBuffer[usAxis].AxisIndex, us_value:=usValue, sd_data:=usPData);
    else
      MyPara.uiCmd    := BUSIF_DRIVEMNGBASE_SET_SYNC_PARA;
      MyPara.aPara[0] := to_dint(AxBuffer[usAxis].AxisIndex);
      MyPara.aPara[1] := to_dint(usValue);
      MyPara.aPara[2] := to_dint(usPData);

      ToBusIF.NewInst(#MyPara, #MyResult);
      retcode := MyResult.aData[0]$DINT;
    end_if;
  else
    retcode := -1;
  end_if;

END_FUNCTION

FUNCTION GLOBAL _DriveMngBase::GetSyncEntry
	VAR_INPUT
		usAxis 	: USINT;
		usValue : USINT;
		usPData : ^DINT;
	END_VAR
	VAR_OUTPUT
		retcode : DINT;
	END_VAR
  VAR
    MyPara   : CmdStruct;
    MyResult : results;
  END_VAR

  if usAxis >= 0 & usAxis < SDDMAXENTRIES then //HasHan
    if bVaranConnected then
      retcode:=toVaran.GetSyncParameter(us_Axis:=AxBuffer[usAxis].AxisIndex, us_value:=usValue, p_data:=usPData);
    else
      MyPara.uiCmd    := BUSIF_DRIVEMNGBASE_GET_SYNC_PARA;
      MyPara.aPara[0] := to_dint(AxBuffer[usAxis].AxisIndex);
      MyPara.aPara[1] := to_dint(usValue);
      MyPara.aPara[2] := (usPData)$DINT;

      ToBusIF.NewInst(#MyPara, #MyResult);
      retcode := MyResult.aData[0]$DINT;
    end_if;
  else
    retcode := -1;
  end_if;

END_FUNCTION

FUNCTION GLOBAL _DriveMngBase::GetDriveType
	VAR_INPUT
		HWCode 	: DINT;
	END_VAR
	VAR_OUTPUT
		DriveType 	: _DRIVETYPE;
	END_VAR
  VAR
  	buffer   : DINT;
    MyPara   : CmdStruct;
    MyResult : results;
    dRetCode : iprStates;
  END_VAR

  //LanSte 27.07.2021 When adding new drivetypes GetDriveTypeStr must also be updated!

  if bVaranConnected then
    buffer := HWCode SHR 16;
    case buffer of
    // 3 Achsen
      0: DriveType:=_SDD_310;
      1: DriveType:=_SDD_315;
      2: DriveType:=_S_340;
      3: DriveType:=_SDD_310;
      4: DriveType:=_S_340;
      6: DriveType:=_SDD_315;
     12: DriveType:=_SDD_335;
     16: DriveType:=_SDD_305;
     20: DriveType:=_SDD_305;
     26: DriveType:=_SDD_310;

     // 2 Achsen
      5: DriveType:=_SDD_215;
      9: DriveType:=_SDD_210;
     22: DriveType:=_SDD_205;

     // 1 Achse
      7: DriveType:=_SDD_120;
     21: DriveType:=_SDD_105;
     10: DriveType:=_SDD_115;

    else
      if DeviceID = DIASDRIVE_MINI_DEVICE_ID then
        DriveType := _MDD_100;
      else
        DriveType:=_NotFound;
      end_if;
    end_case;

  else
    //if businterface is connected
    MyPara.uiCmd    := BUSIF_DRIVEMNGBASE_GET_BUSTYPE;
    //first parameter is the length of followed data
    MyPara.aPara[0] := 0;

    dRetCode := ToBusIF.NewInst(#MyPara, #MyResult);

    if dRetCode = Ready
    & MyResult.uiLng = 1 then
      if MyResult.aData[0] = HWT_ESCAPE_SDIAS then
        case DeviceID of
          DRIVEMNG_BUSDEVICEID_DC061:
            DriveType := _DC061;

          DRIVEMNG_BUSDEVICEID_DC062:
            DriveType := _DC062;

          DRIVEMNG_BUSDEVICEID_SR011:
            DriveType := _SR011;

          DRIVEMNG_BUSDEVICEID_SR012:
            DriveType := _SR012;

          DRIVEMNG_BUSDEVICEID_DC101:
            DriveType := _DC101;

          DRIVEMNG_BUSDEVICEID_DC102:
            DriveType := _DC102;

        else
          DriveType:=_NotFound;
        end_case;

      elsif MyResult.aData[0] = HWT_ESCAPE_VARAN then
        case DeviceID of
          DRIVEMNG_BUSDEVICEID_SDD1300:
            DriveType := _SDD_1300;

          DRIVEMNG_BUSDEVICEID_SDD1400:
            DriveType := _SDD_1400;

          DRIVEMNG_BUSDEVICEID_SDD1500:
            DriveType := _SDD_1500;

          DRIVEMNG_BUSDEVICEID_SDD1600:
            DriveType := _SDD_1600;

          DRIVEMNG_BUSDEVICEID_VSDC151:

            //Check I-Type to display correct Drive type (both VSDC151 and VSDC152 have the same Varan device ID but different I-TYPE parameter values)
            if Parameter_I_Type = DRIVEMNG_I_TYPE_VSDC151 then
              DriveType := _VSDC_151;
            elsif Parameter_I_Type = DRIVEMNG_I_TYPE_VSDC152 then
              DriveType := _VSDC_152;
            else
              DriveType:=_NotFound;
            end_if;

          DRIVEMNG_BUSDEVICEID_MDD2000:
            DriveType := _MDD_2000;

        else
          DriveType:=_NotFound;

        end_case;

      elsif MyResult.aData[0] = HWT_ESCAPE_VARAN_S2 then
        case DeviceID of

          DRIVEMNG_BUSDEVICEID_WA011:
            DriveType := _WA011;

          DRIVEMNG_BUSDEVICEID_WA012:
            DriveType := _WA012;

        else
          DriveType:=_NotFound;

        end_case;

      else
        DriveType:=_NotFound;
      end_if;

    else
      DriveType:=_NotFound;
    end_if;
  end_if;

END_FUNCTION

FUNCTION GLOBAL _DriveMngBase::GetVaranDriveState
	VAR_OUTPUT
		retcode 	: DINT;
	END_VAR
  VAR
    MyPara   : CmdStruct;
    MyResult : results;
  END_VAR

  if bVaranConnected then
    retcode := toVaran.GetDriveIntState();
  else
    MyPara.uiCmd := BUSIF_DRIVEMNGBASE_GET_DRIVE_INT_STATE;
    ToBusIF.NewInst(#MyPara, #MyResult);
    retcode := MyResult.aData[0]$DINT;
  end_if;

END_FUNCTION

FUNCTION GLOBAL _DriveMngBase::SetTimeBase
	VAR_INPUT
		ud_timebase_ms 	: UDINT;
	END_VAR
	VAR_OUTPUT
		sd_retval 	: DINT;
	END_VAR

  //When the DriveMng is called manuelly instead of setting the CyWork Time,
  //the Customer has to tell the Class, witch TimeBase is set, because this Time is use somewhere in the Class.

  IF InitCounter <= 1 THEN  //The Init use the ud_TimeoutCycles and set any value, to prevent
                            //the override from this Value after the Customer has set the TimeBase manuelly, this Methode only works after the first Init run.
    sd_retval := -1;
  else
    IF ud_timebase_ms <> 0 THEN
      ud_timebase_ms *= 1000; // Rev. 1.16: us is the unit for the calculation
      udCycleTimems := ud_timebase_ms;  //save for timeout calculation
      ud_TimeoutCycles := ( SDD_ASY_TIMEOUT / ud_timebase_ms ) + 5;
      sd_retval := 0;
    ELSE
      sd_retval := -2;
    END_IF;
  END_IF;

END_FUNCTION

FUNCTION _DriveMngBase::_DriveMngBase
	VAR_OUTPUT
		ret_code 	: ConfStates;
	END_VAR

  //Rev. 1.16: to avoid wrong information on server if drive is used as a transparent client
  CmdState := _NotInitialized;

  ret_code := C_OK;

END_FUNCTION

FUNCTION VIRTUAL _DriveMngBase::GetBusDeviceID
	VAR_OUTPUT
		output 	: UDINT;
	END_VAR

  //Overwrite this method in derived class
  output := HWC_INVALID_DEVICE_ID;

END_FUNCTION

FUNCTION VIRTUAL _DriveMngBase::GetDrvDeviceID
	VAR_OUTPUT
		output 	: UDINT;
	END_VAR

  //Overwrite this method in derived class
  output := HWC_INVALID_DEVICE_ID;

END_FUNCTION

FUNCTION GLOBAL _DriveMngBase::IsAnyAxisEnabled
	VAR_OUTPUT
		AnyAxisEnabled 	: BOOL;
	END_VAR
  VAR
    UserPara     : CmdStruct;
    UserResult   : Results;
    x            : USINT;
    pThisNewInst : ^void;
  END_VAR

  // search for any enabled axis (all axis must be disabled to set absolut position, because drive needs to switch communication)
  AnyAxisEnabled := FALSE;
  UserPara.uiCmd := SDD_GET_ANY_AXIS_ENABLED;

  for x := 0 to (SDDMAXENTRIES - 1) do
    if (AxBuffer[x].pThis <> NIL) then
      if (AxBuffer[x].AxisOk = 1) then
        UserResult.uiLng := 0;

        pThisNewInst := AxBuffer[x].pThis;
        pThisNewInst$^VirtualBase^.NewInst(#UserPara, #UserResult);

        // if there is an enabled axis
        if (UserResult.uiLng = 1) & UserResult.aData[0] then
          // leave method
          AnyAxisEnabled := TRUE;
          return;
        end_if;
      end_if;
    end_if;
  end_for;

END_FUNCTION

FUNCTION GLOBAL _DriveMngBase::DisableDevice
	VAR_OUTPUT
		RetCode 	: DINT;
	END_VAR
  VAR
    MyPara   : CmdStruct;
    MyResult : results;
  END_VAR

  if bVaranConnected then
    RetCode := toVaran.DisableDevice();
  else
    MyPara.uiCmd    := BUSIF_DRIVEMNGBASE_WRITE_PARAMETER;
    Mypara.aPara[0] := _BUS_IF_DRVMNG_DISABLE_DEVICE;
    RetCode$UDINT   := ToBusIF.NewInst(#MyPara, #MyResult);
    if RetCode$IprStates = ERROR then
      RetCode := -1;
    end_if;
  end_if;

END_FUNCTION

FUNCTION GLOBAL _DriveMngBase::EnableDevice
	VAR_OUTPUT
		RetCode 	: DINT;
	END_VAR
  VAR
    MyPara   : CmdStruct;
    MyResult : results;
  END_VAR

  if bVaranConnected then
    RetCode := toVaran.EnableDevice();
  else
    MyPara.uiCmd    := BUSIF_DRIVEMNGBASE_WRITE_PARAMETER;
    Mypara.aPara[0] := _BUS_IF_DRVMNG_ENABLE_DEVICE;
    RetCode$UDINT   := ToBusIF.NewInst(#MyPara, #MyResult);
    if RetCode$IprStates = ERROR then
      RetCode := -1;
    end_if;
  end_if;

END_FUNCTION

FUNCTION VIRTUAL GLOBAL _DriveMngBase::GetDriveTypeStr
	VAR_INPUT
		eDriveType 	: _DRIVETYPE;
		pDriveTypeStr 	: ^CHAR;
    DriveTypeStrSize : UDINT;
	END_VAR
  VAR
  	tmpstr : array [0..20] of char;
  END_VAR

  if pDriveTypeStr then

    case eDriveType of
      _DRIVETYPE::_NotFound:
        _strcpy(dest:=#tmpstr[0], src:="DiasDrive");
      _DRIVETYPE::_SDD_310:
        _strcpy(dest:=#tmpstr[0], src:="SDD310");
      _DRIVETYPE::_SDD_315:
        _strcpy(dest:=#tmpstr[0], src:="SDD315");
      _DRIVETYPE::_SDD_105:
        _strcpy(dest:=#tmpstr[0], src:="SDD105");
      _DRIVETYPE::_SDD_120:
        _strcpy(dest:=#tmpstr[0], src:="SDD120");
      _DRIVETYPE::_SDD_305:
        _strcpy(dest:=#tmpstr[0], src:="SDD305");
      _DRIVETYPE::_SDD_335:
        _strcpy(dest:=#tmpstr[0], src:="SDD335");
      _DRIVETYPE::_SDD_215:
        _strcpy(dest:=#tmpstr[0], src:="SDD215");
      _DRIVETYPE::_SDD_205:
        _strcpy(dest:=#tmpstr[0], src:="SDD205");
      _DRIVETYPE::_SDD_210:
        _strcpy(dest:=#tmpstr[0], src:="SDD210");
      _DRIVETYPE::_MDD_100:
        _strcpy(dest:=#tmpstr[0], src:="MDD100");
      _DRIVETYPE::_S_340: // ?
        _strcpy(dest:=#tmpstr[0], src:="DiasDrive");
      _DRIVETYPE::_SDD_115:
        _strcpy(dest:=#tmpstr[0], src:="SDD115");
      _DRIVETYPE::_SDD_1300:
        _strcpy(dest:=#tmpstr[0], src:="SDD1300");
      _DRIVETYPE::_SDD_1400:
        _strcpy(dest:=#tmpstr[0], src:="SDD1400");
      _DRIVETYPE::_SDD_1500:
        _strcpy(dest:=#tmpstr[0], src:="SDD1500");
      _DRIVETYPE::_SDD_1600:
        _strcpy(dest:=#tmpstr[0], src:="SDD1600");
      _DRIVETYPE::_MDD_2000:
        _strcpy(dest:=#tmpstr[0], src:="MDD2000");
  	  _DRIVETYPE::_VSDC_151:
        _strcpy(dest:=#tmpstr[0], src:="VSDC151");
  	  _DRIVETYPE::_VSDC_152:
        _strcpy(dest:=#tmpstr[0], src:="VSDC152");
      _DRIVETYPE::_DC061:
        _strcpy(dest:=#tmpstr[0], src:="DC061");
      _DRIVETYPE::_DC062:
        _strcpy(dest:=#tmpstr[0], src:="DC062");
      _DRIVETYPE::_SR011:
        _strcpy(dest:=#tmpstr[0], src:="SR011");
      _DRIVETYPE::_SR012:
        _strcpy(dest:=#tmpstr[0], src:="SR012");
      _DRIVETYPE::_DC101:
        _strcpy(dest:=#tmpstr[0], src:="DC101");
      _DRIVETYPE::_DC102:
        _strcpy(dest:=#tmpstr[0], src:="DC102");
      _DRIVETYPE::_WA011:
        _strcpy(dest:=#tmpstr[0], src:="WA011");
      _DRIVETYPE::_WA012:
        _strcpy(dest:=#tmpstr[0], src:="WA012");
      else
        _strcpy(dest:=#tmpstr[0], src:="DiasDrive");
    end_case;

    if (_strlen(src:=#tmpstr[0]) + 1) <= DriveTypeStrSize then  // +1 for 0 termination
      _strcpy(dest:=pDriveTypeStr, src:=#tmpstr[0] );
    end_if;

  end_if;

END_FUNCTION

FUNCTION VIRTUAL _DriveMngBase::GetSystemTime

  sigclib_getsysdate(pdate:=#sTimeVars.tSysDate);
  sigclib_getsystime(ptime:=#sTimeVars.tSysTime);

  //check for not set time stamp
  if sTimeVars.tSysDate.wYear < 2000 then
    sTimeVars.tSysDate.wYear := 2000;
  end_if;

  //YEAR     MONTH      DAY      HOUR    MINUTE     SEC
  //31 26    25 22     21 17    16 12    11   6    5  0
  //  3F       0F        1F       1F       3F       3F

  //set time and date with structure from drive firmware
  sTimeVars.hdKDATEP241 := sTimeVars.tSysTime.wSecond
                           OR (sTimeVars.tSysTime.wMinute shl 6)
                           OR (sTimeVars.tSysTime.wHour shl 12)
                           OR (sTimeVars.tSysDate.wDay shl 17)
                           OR (sTimeVars.tSysDate.wMonth shl 22)
                           OR ((sTimeVars.tSysDate.wYear-2000) shl 26);

END_FUNCTION

FUNCTION VIRTUAL _DriveMngBase::SetSystemTimeAtDrive
	VAR_INPUT
		AxisNo 	: USINT;
	END_VAR

  //Method is called only in derivations when it is needed to set the sysdate/time to the drive firmware (e.g MDD2000 or VSDC151)

  if sTimeVars.bTimeIsSet = FALSE
  & ((ops.tAbsolute-sTimeVars.udLastWrite) >= DRIVEMNG_WRITE_PLCTIME) | (sTimeVars.udLastWrite = 0) then      //check if time is 0 to write time at startup once

    //get System Time
    GetSystemTime();

    //set system time and date at drive
    if AddASyncEntryDS402( AxisNo       :=  AxisNo
                         , uiParaID     :=  0xFFFF
                         , usParaSubID  :=  SDD_K_DATE
                         , usRdWr       :=  TRUE
                         , pValue       :=  (#sTimeVars.hdKDATEP241)$^USINT
                         , bsDataInfo   :=  0
                         , pThisObj     :=  this
                         , usEntry      :=  0
                         ) = 0 then

      // time is set at drive, store timestamp for next time update
      sTimeVars.udLastWrite := ops.tAbsolute - sigclib_random(DRIVEMNG_SDO_TIMOUT);
    end_if;
  end_if;

END_FUNCTION

FUNCTION VIRTUAL GLOBAL _DriveMngBase::GetFile
	VAR_INPUT
		pDestinationDPNE 	: ^CHAR;
		pFileNameDrive 	: ^CHAR;
		pFilePathDrive 	: ^CHAR;
		pdError 	: ^DINT;(* := nil *)
	END_VAR
	VAR_OUTPUT
		retcode 	: iprStates;
	END_VAR
  VAR
    MyPara   : CmdStruct;
    MyResult : results;
  END_VAR

  retcode := CheckFileHandlingAvailable(pdError);

  if retcode = READY then

    MyPara.uiCmd    := BUSIF_DRIVEMNGBASE_GET_FILE;
    MyPara.aPara[0] := BUSIF_DRIVEMNGBASE_GET_FILE_CB_VER1$DINT;  //Version
    MyPara.aPara[1] := pDestinationDPNE$DINT;
    MyPara.aPara[2] := pFileNameDrive$DINT;
    MyPara.aPara[3] := pFilePathDrive$DINT;
    MyPara.aPara[4] := pdError$DINT;

    retcode := ToBusIF.NewInst(#MyPara, #MyResult);

    if retcode <> READY then
      // Failed to start filehandling, release lock
      ReleaseFileHandling();

      // Set ErrorCode if not already set in NewInst
      if pdError & (pdError^ = DRIVEMNG_FILE_HANDLING_RETCODE_NOERROR) then
        pdError^ := DRIVEMNG_FILE_HANDLING_RETCODE_NOT_SUPPORTED;
      end_if;

#ifdef DEBUG_DRIVEMNGBASE
      if retcode <> ERROR then
        // Unreachable Code
        ((0)$^USINT)^ := 0;
      end_if;
#endif
    end_if;

  end_if;

END_FUNCTION

FUNCTION VIRTUAL GLOBAL _DriveMngBase::GetLogFile
	VAR_INPUT
		pDestinationDPNE 	: ^CHAR;(* := NIL *)
		pdError 	: ^DINT;(* := nil *)
		udFileSelectID 	: UDINT;(* := DRIVEMNG_FILESELECT_LOGFILE *)
	END_VAR
	VAR_OUTPUT
		retcode 	: iprStates;
	END_VAR

  retcode := CheckFileHandlingAvailable(pdError, DRIVEMNG_FILE_RESERVE_IDGETLOGFILE);

  if retcode = READY then

    if pDestinationDPNE then
      // Safe Destination File
      _strcpy(dest:=#s_LogFileV.aDestinationLogFile[0], src:=pDestinationDPNE);
    else
      // Clear Destination File
      s_LogFileV.aDestinationLogFile[0] := 0;  // 0 Termination
    end_if;

    s_LogFileV.udFileSelectId := udFileSelectID;

    s_LogFileV.eGetLogFileSSW := StartGetLogFileSSW;

  end_if;

END_FUNCTION

FUNCTION VIRTUAL GLOBAL _DriveMngBase::GetFileState
	VAR_INPUT
		pdError 	: ^DINT;(* := nil *)
		pdProgress 	: ^DINT;(* := nil *)
		pudBytesRead 	: ^UDINT;(* := nil *)
	END_VAR
	VAR_OUTPUT
		retcode 	: iprStates;
	END_VAR
  VAR
    MyPara   : CmdStruct;
    MyResult : results;
  END_VAR

  if bVaranConnected then
    retcode := ERROR; //Not supported with _VaranDriveBase class
    if pdError then
      pdError^:= DRIVEMNG_FILE_HANDLING_RETCODE_NOT_SUPPORTED;
    end_if;
  else

    if Online.read() = 0 then
      retcode := ERROR; //Drive is not online
      if pdError then
        pdError^ := DRIVEMNG_FILE_HANDLING_RETCODE_NOT_ONLINE;
      end_if;
      return;
    end_if;

    // Check if filehandling is active only in busif
    if (sigclib_atomic_getU32(pValue:=#ud_FileHandlingReserved) = DRIVEMNG_FILE_RESERVE_IDDEFAULT) then

      // Pass on command to Busif
      MyPara.uiCmd    := BUSIF_DRIVEMNGBASE_GET_FILE_STATE;
      MyPara.aPara[0] := BUSIF_DRIVEMNGBASE_GET_FILE_STATE_CB_VER1$DINT;  //Version
      MyPara.aPara[1] := pdError$DINT;
      MyPara.aPara[2] := pdProgress$DINT;
      MyPara.aPara[3] := pudBytesRead$DINT;

      retcode := ToBusIF.NewInst(#MyPara, #MyResult);

      if (retcode = READY) | (retcode = ERROR) then
        // File handling has completed => unlock
        ReleaseFileHandling();
      end_if;

    // Check if filehandling is active get log file
    elsif (sigclib_atomic_getU32(pValue:=#ud_FileHandlingReserved) = DRIVEMNG_FILE_RESERVE_IDGETLOGFILE) then

      if s_LogFileV.eGetLogFileSSW = wait4GetLogFile then

        // Pass on command to Busif
        MyPara.uiCmd    := BUSIF_DRIVEMNGBASE_GET_FILE_STATE;
        MyPara.aPara[0] := BUSIF_DRIVEMNGBASE_GET_FILE_STATE_CB_VER1$DINT;  //Version
        MyPara.aPara[1] := pdError$DINT;
        MyPara.aPara[2] := pdProgress$DINT;
        MyPara.aPara[3] := pudBytesRead$DINT;

        retcode := ToBusIF.NewInst(#MyPara, #MyResult);

        if (retcode = READY) | (retcode = ERROR) then
          // Reset SSW
          s_LogFileV.eGetLogFileSSW := IdleGetLogFile;
          // File handling has completed => unlock
          ReleaseFileHandling();
        end_if;

      elsif s_LogFileV.eGetLogFileSSW = ErrorGetLogFile then

        retcode := ERROR;

        if pdError then
          pdError^ := s_LogFileV.ErrorCodeLogFile;
        end_if;

        s_LogFileV.eGetLogFileSSW := IdleGetLogFile;

        // File handling has completed => unlock
        ReleaseFileHandling();

      elsif s_LogFileV.eGetLogFileSSW = IdleGetLogFile then

#ifdef DEBUG_DRIVEMNGBASE
        // Unreachable Code
        #pragma message("LanSte 02.06.2022 12:43 \ TODO Remove for release Version")
        ((0)$^USINT)^ := 0;
#endif

        retcode := READY;
        ReleaseFileHandling();

      else

        // Busy in SSW
        retcode := BUSY;

        if pdError then
          pdError^ := DRIVEMNG_FILE_HANDLING_RETCODE_NOERROR;
        end_if;

      end_if;

    else

      // No File handling active, ready for new.
      retcode := READY;
      if pdError then
        pdError^ := DRIVEMNG_FILE_HANDLING_RETCODE_NOERROR;
      end_if;

    end_if;

  end_if;

END_FUNCTION

FUNCTION VIRTUAL GLOBAL _DriveMngBase::SetFile
	VAR_INPUT
		pWriteData 	: ^void;
		udWriteDataLen 	: UDINT;
		pFilePathDrive 	: ^CHAR;
		pFileNameDrive 	: ^CHAR;
		pdError 	: ^DINT;(* := nil *)
	END_VAR
	VAR_OUTPUT
		retcode 	: iprStates;
	END_VAR
  VAR
    MyPara   : CmdStruct;
    MyResult : results;
  END_VAR

  retcode := CheckFileHandlingAvailable(pdError);

  if retcode = READY then

    //we are connected via businterface
    MyPara.uiCmd    := BUSIF_DRIVEMNGBASE_SET_FILE;
    MyPara.aPara[0] := BUSIF_DRIVEMNGBASE_SET_FILE_CB_VER1$DINT;  //Version
    MyPara.aPara[1] := pWriteData$DINT;
    MyPara.aPara[2] := udWriteDataLen$DINT;
    MyPara.aPara[3] := pFilePathDrive$DINT;
    MyPara.aPara[4] := pFileNameDrive$DINT;
    MyPara.aPara[5] := pdError$DINT;

    retcode := ToBusIF.NewInst(#MyPara, #MyResult);

    if retcode <> READY then
      // Failed to start filehandling, release lock
      ReleaseFileHandling();

      // Set ErrorCode if not already set in NewInst
      if pdError & (pdError^ = DRIVEMNG_FILE_HANDLING_RETCODE_NOERROR) then
        pdError^ := DRIVEMNG_FILE_HANDLING_RETCODE_NOT_SUPPORTED;
      end_if;

#ifdef DEBUG_DRIVEMNGBASE
      if retcode <> ERROR then
        // Unreachable Code
        ((0)$^USINT)^ := 0;
      end_if;
#endif
    end_if;
  end_if;

END_FUNCTION

FUNCTION VIRTUAL GLOBAL _DriveMngBase::GetFileSize
	VAR_INPUT
    pFileNameDrive 	: ^CHAR;
    pFilePathDrive 	: ^CHAR;
    pudSize 	: ^UDINT;
    pdError 	: ^DINT;(* := nil *)
	END_VAR
	VAR_OUTPUT
		retcode 	: iprStates;
	END_VAR
  VAR
    MyPara   : CmdStruct;
    MyResult : results;
  END_VAR

  retcode := CheckFileHandlingAvailable(pdError);

  if retcode = READY then

    //we are connected via businterface
    MyPara.uiCmd    := BUSIF_DRIVEMNGBASE_GET_FILE_SIZE;
    MyPara.aPara[0] := BUSIF_DRIVEMNGBASE_GET_FILE_SIZE_CB_VER1$DINT;  //Version
    MyPara.aPara[1] := pFileNameDrive$DINT;
    MyPara.aPara[2] := pFilePathDrive$DINT;
    MyPara.aPara[3] := pudSize$DINT;
    MyPara.aPara[4] := pdError$DINT;

    retcode := ToBusIF.NewInst(#MyPara, #MyResult);

    if retcode <> READY then
      // Failed to start filehandling, release lock
      ReleaseFileHandling();

      // Set ErrorCode if not already set in NewInst
      if pdError & (pdError^ = DRIVEMNG_FILE_HANDLING_RETCODE_NOERROR) then
        pdError^ := DRIVEMNG_FILE_HANDLING_RETCODE_NOT_SUPPORTED;
      end_if;

#ifdef DEBUG_DRIVEMNGBASE
      if retcode <> ERROR then
        // Unreachable Code
        ((0)$^USINT)^ := 0;
      end_if;
#endif
    end_if;
  end_if;

END_FUNCTION

FUNCTION VIRTUAL GLOBAL _DriveMngBase::GetFileBuffer
	VAR_INPUT
		pFileNameDrive 	: ^CHAR;
		pFilePathDrive 	: ^CHAR;
		udBufferSize 	: UDINT;
		pDataBuffer 	: ^void;(* := nil *)
		udDataLenToRead 	: UDINT;(* := 0 *)
		pdError 	: ^DINT;(* := nil *)
	END_VAR
	VAR_OUTPUT
		retcode 	: iprStates;
	END_VAR
  VAR
    MyPara   : CmdStruct;
    MyResult : results;
  END_VAR

  retcode := CheckFileHandlingAvailable(pdError);

  if retcode = READY then

    //we are connected via businterface
    MyPara.uiCmd    := BUSIF_DRIVEMNGBASE_GET_FILE_BUFFER;
    MyPara.aPara[0] := BUSIF_DRIVEMNGBASE_GET_FILE_BUFFER_CB_VER1$DINT;  //Version
    MyPara.aPara[1] := pFileNameDrive$DINT;
    MyPara.aPara[2] := pFilePathDrive$DINT;
    MyPara.aPara[3] := udBufferSize$DINT;
    MyPara.aPara[4] := pDataBuffer$DINT;
    MyPara.aPara[5] := udDataLenToRead$DINT;
    MyPara.aPara[6] := pdError$DINT;

    retcode := ToBusIF.NewInst(#MyPara, #MyResult);

    if retcode <> READY then
      // Failed to start filehandling, release lock
      ReleaseFileHandling();

      // Set ErrorCode if not already set in NewInst
      if pdError & (pdError^ = DRIVEMNG_FILE_HANDLING_RETCODE_NOERROR) then
        pdError^ := DRIVEMNG_FILE_HANDLING_RETCODE_NOT_SUPPORTED;
      end_if;
#ifdef DEBUG_DRIVEMNGBASE
      if retcode <> ERROR then
        // Unreachable Code
        ((0)$^USINT)^ := 0;
      end_if;
#endif
    end_if;
  end_if;

END_FUNCTION

FUNCTION VIRTUAL _DriveMngBase::GetLogFileCyclic
  VAR
    retcode  : iprStates;
    MyPara   : CmdStruct;
    MyResult : results;
    aFileNameDrive    : ARRAY [0..199] OF CHAR;
    aFilePathDrive    : ARRAY [0..199] OF CHAR;
    usAxisNo : USINT;
  END_VAR

  case s_LogFileV.eGetLogFileSSW of

//*****************************************************************************
    t_e_GetLogFileSSW::IdleGetLogFile:
      // Do Nothing

//*****************************************************************************
    t_e_GetLogFileSSW::StartGetLogFileSSW,
    t_e_GetLogFileSSW::WriteLOGFileParam:

      s_LogFileV.ErrorCodeLogFile := DRIVEMNG_FILE_HANDLING_RETCODE_NOERROR;  // Fehlercode zurücksetzen

      //Only allow to get logfile if no axis is enabled
      if IsAnyAxisEnabled() = FALSE then

        // get the standard information of the drive
        usAxisNo := GetFirstAxIndex();

        if usAxisNo <> 16#FF then
          //We have to tell the firmware that the logfile should be written

          //Writing to K-LOG leads to that the firmware is going to write their logbuffer into the logfile on the drive
          //This will block the other asynchronous communication and can take some seconds
          //Give this access a high timeout so we won't get an error with the default timeout

          // Get usParaLogIdx and dParaLogVal from derived class
          GetLogFileWrParam(pParaIDX:=#s_LogFileV.usParaLogIdx, pParaVal:=#s_LogFileV.dParaLogVal, pParaTimeout:=#s_LogFileV.udParaLogTimeout,s_LogFileV.udFileSelectId);

          if s_LogFileV.usParaLogIdx then
            if AddASyncEntry(AxisNo    :=  usAxisNo
                           , usParaNr  :=  s_LogFileV.usParaLogIdx
                           , usRdWr    :=  1
                           , dValue    :=  s_LogFileV.dParaLogVal  //Start to write logfile
                           , pThisObj  :=  this
                           , usEntry   :=  0
                           , udTimeout :=  s_LogFileV.udParaLogTimeout) = 0 then

              s_LogFileV.bWait4LogFilePara := TRUE;
              s_LogFileV.udTimeStampLogPara := ops.tAbsolute;
              s_LogFileV.eGetLogFileSSW := t_e_GetLogFileSSW::Wait4WrLOGFileResponse;
            end_if;
          else
            // usParaLogIdx not used to write parameter, skip step.
            s_LogFileV.eGetLogFileSSW := t_e_GetLogFileSSW::ReadLOGFileParam;
          end_if;

        else

          s_LogFileV.ErrorCodeLogFile := DRIVEMNG_FILE_HANDLING_RETCODE_NOT_ONLINE;  //Drive is not online
          s_LogFileV.eGetLogFileSSW := t_e_GetLogFileSSW::ErrorGetLogFile;

        end_if;
      else

        s_LogFileV.ErrorCodeLogFile := DRIVEMNG_FILE_HANDLING_RETCODE_AXIS_ENABLED;  //Axis must be not enabled to start get logfile
        s_LogFileV.eGetLogFileSSW := t_e_GetLogFileSSW::ErrorGetLogFile;

      end_if;

//*****************************************************************************
    t_e_GetLogFileSSW::Wait4WrLOGFileResponse:
      //Wait until we get response from K_LOG
      if s_LogFileV.bWait4LogFilePara = FALSE then

        // Check Return Value
        if s_LogFileV.dParaLogValRd <> 16#7FFFFFFF then
          s_LogFileV.eGetLogFileSSW := t_e_GetLogFileSSW::ReadLOGFileParam;
        else
          s_LogFileV.ErrorCodeLogFile := DRIVEMNG_FILE_HANDLING_RETCODE_WRITEPARA_FAILED;  // Unexpected Para Val was returned
          s_LogFileV.eGetLogFileSSW := t_e_GetLogFileSSW::ErrorGetLogFile;
        end_if;

      elsif ops.tAbsolute - s_LogFileV.udTimeStampLogPara > s_LogFileV.udParaLogTimeout then  //Timeout while waiting for response of K-LOG
        s_LogFileV.ErrorCodeLogFile := DRIVEMNG_FILE_HANDLING_RETCODE_WRITEPARA_TIMEOUT;  // Unexpected Para Val was returned
        s_LogFileV.eGetLogFileSSW := t_e_GetLogFileSSW::ErrorGetLogFile;
      end_if;

//*****************************************************************************
    t_e_GetLogFileSSW::ReadLOGFileParam:

      //Only allow to get logfile if no axis is enabled
      if IsAnyAxisEnabled() = FALSE then

        // get the standard information of the drive
        usAxisNo := GetFirstAxIndex();

        if usAxisNo <> 16#FF then

          // Read back parameters to see if file was successfully copied to drive

          // Get usParaLogIdx and dParaLogVal from derived class
          GetLogFileRdParam(pParaIDX:=#s_LogFileV.usParaLogIdx, pParaVal:=#s_LogFileV.dParaLogVal, pParaTimeout:=#s_LogFileV.udParaLogTimeout,s_LogFileV.udFileSelectId);

          if s_LogFileV.usParaLogIdx then
            if AddASyncEntry(AxisNo    :=  usAxisNo
                           , usParaNr  :=  s_LogFileV.usParaLogIdx
                           , usRdWr    :=  0
                           , dValue    :=  s_LogFileV.dParaLogVal  //Start to write logfile
                           , pThisObj  :=  this
                           , usEntry   :=  0
                           , udTimeout :=  s_LogFileV.udParaLogTimeout) = 0 then

              s_LogFileV.bWait4LogFilePara := TRUE;
              s_LogFileV.udTimeStampLogPara := ops.tAbsolute;
              s_LogFileV.eGetLogFileSSW := t_e_GetLogFileSSW::Wait4RdLOGFileResponse;
            end_if;

          else
            // usParaLogIdx not used to write parameter, skip step.
            s_LogFileV.eGetLogFileSSW := t_e_GetLogFileSSW::StartGetLogFile;
          end_if;

        else

          s_LogFileV.ErrorCodeLogFile := DRIVEMNG_FILE_HANDLING_RETCODE_NOT_ONLINE;  //Drive is not online
          s_LogFileV.eGetLogFileSSW := t_e_GetLogFileSSW::ErrorGetLogFile;

        end_if;
      else

        s_LogFileV.ErrorCodeLogFile := DRIVEMNG_FILE_HANDLING_RETCODE_AXIS_ENABLED;  //Axis must be not enabled to start get logfile
        s_LogFileV.eGetLogFileSSW := t_e_GetLogFileSSW::ErrorGetLogFile;

      end_if;

//*****************************************************************************
    t_e_GetLogFileSSW::Wait4RdLOGFileResponse:
      //Wait until we get response from K_LOG
      if s_LogFileV.bWait4LogFilePara = FALSE then

        // Check Return Value
        if s_LogFileV.dParaLogVal = s_LogFileV.dParaLogValRd then
          s_LogFileV.eGetLogFileSSW := t_e_GetLogFileSSW::StartGetLogFile;
        else
          s_LogFileV.ErrorCodeLogFile := DRIVEMNG_FILE_HANDLING_RETCODE_READBACKPARA_FAILED;  // Unexpected Para Val was returned
          s_LogFileV.eGetLogFileSSW := t_e_GetLogFileSSW::ErrorGetLogFile;
        end_if;

      elsif ops.tAbsolute - s_LogFileV.udTimeStampLogPara > s_LogFileV.udParaLogTimeout then  //Timeout while waiting for response of K-LOG
        s_LogFileV.ErrorCodeLogFile := DRIVEMNG_FILE_HANDLING_RETCODE_READBACKPARA_TIMEOUT;  // Unexpected Para Val was returned
        s_LogFileV.eGetLogFileSSW := t_e_GetLogFileSSW::ErrorGetLogFile;
      end_if;

//*****************************************************************************
    t_e_GetLogFileSSW::StartGetLogFile:
      //Check if user wants to set a specific name or if we should use the default name
      if _strlen(src:=#s_LogFileV.aDestinationLogFile[0]) = 0 then
        GetDefaultLogFileDestinationDPNE(#s_LogFileV.aDestinationLogFile[0], s_LogFileV.udFileSelectId);  //Use default DPNE
      // else
        //Use given DPNE
      end_if;

      GetDefaultLogFileNameDrive(#aFileNameDrive[0],s_LogFileV.udFileSelectId);
      GetDefaultLogFilePathDrive(#aFilePathDrive[0],s_LogFileV.udFileSelectId);

      MyPara.uiCmd    := BUSIF_DRIVEMNGBASE_GET_FILE;
      MyPara.aPara[0] := BUSIF_DRIVEMNGBASE_GET_FILE_CB_VER1$DINT;  //Version
      MyPara.aPara[1] := (#s_LogFileV.aDestinationLogFile[0])$DINT;
      MyPara.aPara[2] := (#aFileNameDrive[0])$DINT;
      MyPara.aPara[3] := (#aFilePathDrive[0])$DINT;
      MyPara.aPara[4] := (#s_LogFileV.ErrorCodeLogFile)$DINT;

      retcode := ToBusIF.NewInst(#MyPara, #MyResult);

      if retcode = READY then
        s_LogFileV.eGetLogFileSSW := t_e_GetLogFileSSW::wait4GetLogFile;
      elsif retcode = ERROR then

        // Check if Error code was set
        if s_LogFileV.ErrorCodeLogFile = DRIVEMNG_FILE_HANDLING_RETCODE_NOERROR then
          s_LogFileV.ErrorCodeLogFile := DRIVEMNG_FILE_HANDLING_RETCODE_NOT_SUPPORTED;
        end_if;

        s_LogFileV.eGetLogFileSSW := t_e_GetLogFileSSW::ErrorGetLogFile;
      else
#ifdef DEBUG_DRIVEMNGBASE
        // Unreachable Code
        #pragma message("LanSte 02.06.2022 12:43 \ TODO Remove for release Version")
        ((0)$^USINT)^ := 0;
#endif
      end_if;

//*****************************************************************************
    t_e_GetLogFileSSW::wait4GetLogFile:
      // Wait for User to call GetFileState

//*****************************************************************************
    t_e_GetLogFileSSW::ErrorGetLogFile:
      // Wait for User to call GetFileState

  end_case;

END_FUNCTION

FUNCTION VIRTUAL _DriveMngBase::GetLogFileWrParam
	VAR_INPUT
		pParaIDX 	: ^USINT;
		pParaVal 	: ^DINT;
		pParaTimeout 	: ^UDINT;
		FileSelect 	: UDINT;
	END_VAR

  // Default Implementation, not supported. Override in derived Classes for support
  if pParaIDX then
    pParaIDX^ := 0;
  end_if;

  if pParaVal then
    pParaVal^ := 0;
  end_if;

  if pParaTimeout then
    pParaTimeout^ := DRIVEMNG_FILE_HANDLING_TIMEOUT_LOG_PARAM;
  end_if;

END_FUNCTION

FUNCTION VIRTUAL _DriveMngBase::GetLogFileRdParam
	VAR_INPUT
		pParaIDX 	: ^USINT;
		pParaVal 	: ^DINT;
		pParaTimeout 	: ^UDINT;
		FileSelect 	: UDINT;
	END_VAR

  // Default Implementation, not supported. Override in derived Classes for support
  if pParaIDX then
    pParaIDX^ := 0;
  end_if;

  if pParaVal then
    pParaVal^ := 0;
  end_if;

  if pParaTimeout then
    pParaTimeout^ := DRIVEMNG_FILE_HANDLING_TIMEOUT_LOG_PARAM;
  end_if;

END_FUNCTION

FUNCTION VIRTUAL _DriveMngBase::GetDefaultLogFileDestinationDPNE
	VAR_INPUT
		pDPNE 	: ^CHAR;
		FileSelect 	: UDINT;(* := 0 *)
	END_VAR
  VAR
    aSerialNo         : ARRAY [0..10] OF CHAR;
  END_VAR

  if pDPNE then

    if FileSelect = DRIVEMNG_FILESELECT_DEBUGLOGFILE then
      _strcpy(dest:=pDPNE, src:=DRIVEMNG_DEFAULT_CPU_DEBUGLOGFILENAME_PATH );
    else
      _strcpy(dest:=pDPNE, src:=DRIVEMNG_DEFAULT_CPU_LOGFILENAME_PATH);
    end_if;

    //add serialno as string to filename
    _memset(dest:=#aSerialNo[0], usByte:=0, cntr:=sizeof(aSerialNo));
    sigclib_sprintfST(pd:=#aSerialNo[0], format:="%08d", p0:=#SerialNo);
    _strcat(dest:=pDPNE, src:=#aSerialNo[0]);

    _strcat(dest:=pDPNE, src:=DRIVEMNG_DEFAULT_CPU_LOGFILENAME_EXTENSION);
  end_if;

END_FUNCTION

FUNCTION VIRTUAL _DriveMngBase::GetDefaultLogFileNameDrive
	VAR_INPUT
		pFileName 	: ^CHAR;
		FileSelect 	: UDINT;
	END_VAR

  if pFileName then

    if FileSelect = DRIVEMNG_FILESELECT_DEBUGLOGFILE then
      _strcpy(dest:=pFileName, src:=DRIVEMNG_DEFAULT_DRIVE_DEBUGLOGFILENAME_NAME);
    else
      //Copy default name of Drive logfiles into buffer
      _strcpy(dest:=pFileName, src:=DRIVEMNG_DEFAULT_DRIVE_LOGFILENAME_NAME);
    end_if;

  end_if;

END_FUNCTION

FUNCTION VIRTUAL _DriveMngBase::GetDefaultLogFilePathDrive
	VAR_INPUT
		pFilePath 	: ^CHAR;
		FileSelect 	: UDINT;
	END_VAR

  if pFilePath then
    //Copy default name of Drive logfile path/directory into buffer
    _strcpy(dest:=pFilePath, src:=DRIVEMNG_DEFAULT_DRIVE_LOGFILENAME_PATH);
  end_if;

END_FUNCTION

FUNCTION VIRTUAL _DriveMngBase::CheckFileHandlingAvailable
	VAR_INPUT
		pdError 	: ^DINT;(* := nil *)
		ReserveID 	: UDINT;(* := DRIVEMNG_FILE_RESERVE_IDDEFAULT *)
	END_VAR
	VAR_OUTPUT
		retcode 	: iprStates;
	END_VAR

  // Default
  retcode := ERROR;

  if bVaranConnected then
     //Not supported with _VaranDriveBase class
    if pdError then
      pdError^:= DRIVEMNG_FILE_HANDLING_RETCODE_NOT_SUPPORTED;
    end_if;
  else

    if Online.read() = 0 then
      //Drive is not online
      if pdError then
        pdError^ := DRIVEMNG_FILE_HANDLING_RETCODE_NOT_ONLINE;
      end_if;
      return;
    end_if;

    if ReserveFileHandling(ReserveID) = TRUE then

      retcode := READY;

      // Reset ErrorCode
      if pdError then
        pdError^ := DRIVEMNG_FILE_HANDLING_RETCODE_NOERROR;
      end_if;

    elsif pdError then
      pdError^ := DRIVEMNG_FILE_HANDLING_RETCODE_FILEHANDLING_BUSY;
    end_if;

  end_if;

END_FUNCTION

FUNCTION VIRTUAL _DriveMngBase::ReserveFileHandling
	VAR_INPUT
		ReserveID 	: UDINT;(* := DRIVEMNG_FILE_RESERVE_IDDEFAULT *)
	END_VAR
	VAR_OUTPUT
		bReserverdOK 	: BOOL;
	END_VAR
  VAR
  	ud_FileHandlingReservedOld : UDINT;
  END_VAR

  bReserverdOK := FALSE;

  ud_FileHandlingReservedOld := sigclib_atomic_cmpxchgU32(pValue:=#ud_FileHandlingReserved, cmpVal:=DRIVEMNG_FILE_RESERVE_IDFREE, newVal:=ReserveID);

  if ud_FileHandlingReservedOld = DRIVEMNG_FILE_RESERVE_IDFREE then
    bReserverdOK := TRUE;
  end_if;

END_FUNCTION

FUNCTION VIRTUAL _DriveMngBase::ReleaseFileHandling

  sigclib_atomic_setU32(pValue:=#ud_FileHandlingReserved, value:=DRIVEMNG_FILE_RESERVE_IDFREE); //unlock method

END_FUNCTION
